(* IEC 61131-3 sources: llm-plc-st-eval/data/processed_definitivo/qwen2.5-coder_14b/C4/zero_shot, 3 files *)

(* ---- ejec_1.st ---- *)
FUNCTION_BLOCK FB_D
VAR_INPUT
    demanda : BOOL;  // Indica si hay una demanda de activación de bombas
    falla1 : BOOL;   // Indica si la bomba1 ha fallado
    falla2 : BOOL;   // Indica si la bomba2 ha fallado
END_VAR
VAR_OUTPUT
    bomba1 : BOOL;   // Controla la activación de la bomba1
    bomba2 : BOOL;   // Controla la activación de la bomba2
    almFalla : BOOL; // Almacena la falla detectada
END_VAR
VAR
    turno : BOOL;    // Variable de estado para alternar el turno entre bomba1 y bomba2
    fDem : R_TRIG;   // Detector de flanco de subida en la demanda
END_VAR

// Detecta el flanco de subida en la demanda
fDem(CLK := demanda);

// Si se detecta un flanco de subida en la demanda, se alterna el turno
IF fDem.Q THEN
    turno := NOT turno;
END_IF

// Si hay una demanda de activación de bombas
IF demanda THEN
    // Si es el turno de la bomba1
    IF turno THEN
        bomba1 := NOT falla1;  // Activa bomba1 si no ha fallado
        bomba2 := falla1 AND NOT falla2;  // Activa bomba2 si bomba1 ha fallado y bomba2 no ha fallado
        almFalla := falla1;  // Almacena la falla de bomba1 si ha ocurrido
    // Si es el turno de la bomba2
    ELSE
        bomba2 := NOT falla2;  // Activa bomba2 si no ha fallado
        bomba1 := falla2 AND NOT falla1;  // Activa bomba1 si bomba2 ha fallado y bomba1 no ha fallado
        almFalla := falla2;  // Almacena la falla de bomba2 si ha ocurrido
    END_IF
// Si no hay demanda de activación de bombas
ELSE
    bomba1 := FALSE;  // Desactiva bomba1
    bomba2 := FALSE;  // Desactiva bomba2
    almFalla := FALSE;  // Limpia el registro de falla
END_IF
END_FUNCTION_BLOCK

(* ---- ejec_2.st ---- *)
FUNCTION_BLOCK FB_D
VAR_INPUT
    demanda : BOOL;  // Entrada que indica si hay una demanda de activación de bombas
    falla1 : BOOL;   // Entrada que indica si hay una falla en la bomba 1
    falla2 : BOOL;   // Entrada que indica si hay una falla en la bomba 2
END_VAR
VAR_OUTPUT
    bomba1 : BOOL;   // Salida que controla la activación de la bomba 1
    bomba2 : BOOL;   // Salida que controla la activación de la bomba 2
    almFalla : BOOL; // Salida que indica si hay una falla detectada
END_VAR
VAR
    turno : BOOL;    // Variable interna que controla el turno entre bomba1 y bomba2
    fDem : R_TRIG;   // Objeto de retardo que detecta el flanco de subida de la demanda
END_VAR

// Configuración del objeto de retardo R_TRIG para detectar el flanco de subida de la demanda
fDem(CLK := demanda);

// Si se detecta un flanco de subida en la demanda
IF fDem.Q THEN
    // Cambiar el turno entre bomba1 y bomba2
    turno := NOT turno;
END_IF

// Si hay una demanda de activación de bombas
IF demanda THEN
    // Si el turno está asignado a bomba1
    IF turno THEN
        // Activar bomba1 si no hay falla en bomba1
        bomba1 := NOT falla1;
        // Activar bomba2 si hay falla en bomba1 y no hay falla en bomba2
        bomba2 := falla1 AND NOT falla2;
        // Activar la alarma de falla si hay falla en bomba1
        almFalla := falla1;
    // Si el turno está asignado a bomba2
    ELSE
        // Activar bomba2 si no hay falla en bomba2
        bomba2 := NOT falla2;
        // Activar bomba1 si hay falla en bomba2 y no hay falla en bomba1
        bomba1 := falla2 AND NOT falla1;
        // Activar la alarma de falla si hay falla en bomba2
        almFalla := falla2;
    END_IF
// Si no hay demanda de activación de bombas
ELSE
    // Desactivar bomba1
    bomba1 := FALSE;
    // Desactivar bomba2
    bomba2 := FALSE;
    // Desactivar la alarma de falla
    almFalla := FALSE;
END_IF
END_FUNCTION_BLOCK

(* ---- ejec_3.st ---- *)
FUNCTION_BLOCK FB_D
VAR_INPUT
    demanda : BOOL;  // Indica si hay una demanda de agua
    falla1 : BOOL;   // Indica si la bomba1 ha fallado
    falla2 : BOOL;   // Indica si la bomba2 ha fallado
END_VAR
VAR_OUTPUT
    bomba1 : BOOL;   // Controla el funcionamiento de la bomba1
    bomba2 : BOOL;   // Controla el funcionamiento de la bomba2
    almFalla : BOOL; // Almacena la falla detectada
END_VAR
VAR
    turno : BOOL;    // Variable de estado para alternar entre bombas
    fDem : R_TRIG;   // Temporizador de flanco ascendente para detectar cambios en demanda
END_VAR

// Configura el temporizador de flanco ascendente con la señal de demanda
fDem(CLK := demanda);

// Si hay un flanco ascendente en la demanda
IF fDem.Q THEN
    // Alterna el estado del turno
    turno := NOT turno;
END_IF

// Si hay demanda de agua
IF demanda THEN
    // Si el turno está activo
    IF turno THEN
        // Activa bomba1 si no hay falla en bomba1
        bomba1 := NOT falla1;
        // Activa bomba2 si hay falla en bomba1 y no hay falla en bomba2
        bomba2 := falla1 AND NOT falla2;
        // Almacena la falla de bomba1 si hay falla
        almFalla := falla1;
    ELSE
        // Activa bomba2 si no hay falla en bomba2
        bomba2 := NOT falla2;
        // Activa bomba1 si hay falla en bomba2 y no hay falla en bomba1
        bomba1 := falla2 AND NOT falla1;
        // Almacena la falla de bomba2 si hay falla
        almFalla := falla2;
    END_IF
ELSE
    // Si no hay demanda, apaga ambas bombas
    bomba1 := FALSE;
    bomba2 := FALSE;
    // Limpia el registro de falla
    almFalla := FALSE;
END_IF
END_FUNCTION_BLOCK
